Fanuc KAREL source: ko00071.KL

-- PROVISIONAL review KL for V770-1; original PC SHA256 8d485b9a7683df311446ff979c30c58d440ead07da9b9b3d3b6b09d3f4cb578b
-- Incomplete behavior may be omitted. Consult companion uncertainty JSON. Do not deploy.
PROGRAM KO00071
%NOLOCKGROUP
BEGIN
  -- UNRESOLVED_PC offsets 5-12; opcodes 9D,23
  -- UNRESOLVED_PC offsets 17-66; opcodes 27,22,1C,27,49,7E,AD,22,31,7E,4A
  -- UNRESOLVED_PC offsets 71-75; opcodes 7F
END KO00071
